FUNCTION_BLOCK FB_IEC61850
VAR
	bInitDone: BOOL := FALSE;	

	i: UDINT;
	j: UDINT;
END_VAR

IF NOT bInitDone THEN
	F_IEC61850ServerInit();

	bInitDone := TRUE;
END_IF

FOR i := 1 TO c_nNumTurbines DO
	fbServer[i].Execute();
	FOR j := 1 TO c_nNumSessions DO
		fbSession[i,j]();
	END_FOR
END_FOR

END_FUNCTION_BLOCK

(* stored: Version 1.1.0.1
   POU FB_IEC61850: Id {c4980344-d71e-4ccf-9e09-bede6b67863a}, SpecialFunc None *)
